{attribute 'qualified_only'}
{attribute 'strict'}
{attribute 'to_string'}
TYPE E_Int :
(
	eOptionA := 0,
	eOptionB,
	eOptionC
) INT;
END_TYPE

(* stored: Version 1.1.0.1, ProductVersion 3.1.4026.19
   DUT E_Int: Id {06c73e96-77d3-4a54-8a2d-a71c97362de6} *)
